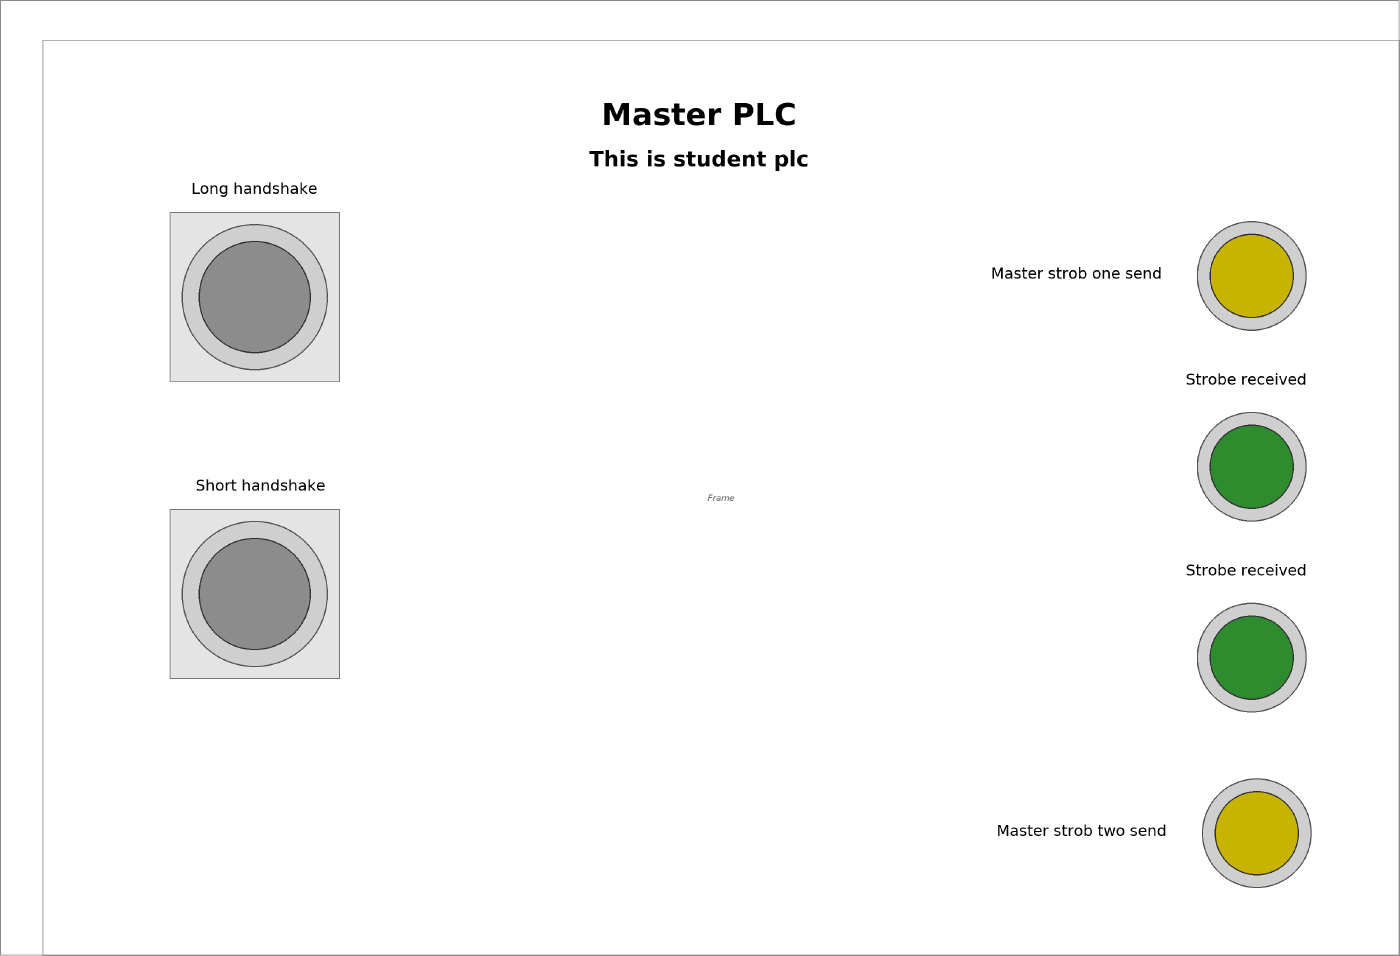
VISUALIZATION VisualizationStudent  // 1650x1127
    Frame (50,47 1600x1080)
    Label (699,110 250x50), "Master PLC"
    PushSwitch (200,250 200x200), variable: GVLStudent.IXButtonLong, behaviour: TAP, style: Switch-PushSwitch-Gray
    PushSwitch (200,600 200x200), variable: GVLStudent.IXButtonShort, behaviour: TAP, style: Switch-PushSwitch-Gray
    Label (225,200 150x45), "Long handshake"
    Label (225,550 164x45), "Short handshake"
    Label (1095,300 348x45), "Master strob one send"
    Lamp1 (1400,475 150x150), variable: GVLStudent.OXLampIXOneGreen, style: Lamp-Lamp1-Green
    Lamp1 (1406,907 150x150), variable: GVLStudent.OXLampOXTwo, style: Lamp-Lamp1-Yellow
    Lamp1 (1400,250 150x150), variable: GVLStudent.OXLampOXOne, style: Lamp-Lamp1-Yellow
    Label (1350,425 238x45), "Strobe received"
    Label (1101,957 348x45), "Master strob two send"
    Lamp1 (1400,700 150x150), variable: GVLStudent.OXLampIXTwoGreen, style: Lamp-Lamp1-Green
    Label (1350,650 238x45), "Strobe received"
    Label (643,172 362x30), "This is student plc"
END_VISUALIZATION

(* stored: Version 1.1.0.1, ProductVersion 3.1.4024.12
   Visu VisualizationStudent: Id {5276086c-0119-418b-ae8f-5e465a97ae16} *)
